SUBAPPLICATION AR_M2M_Subscribe_TO_Q_OPC (* Remote-Subscribe eines fertigen physikalischen Werts (M2M) -> VT-Anzeige (Q_NumericValue_PHYSA, gedrosselt) + VALUE_OUT. Wie AR_M2M_Subscribe_TO_Q_Publish_OPC, aber ohne lokalen Re-Publish. *)
  (* Standard: 61499-2; Description: Copyright (c) 2026 Meisterschulen am Ostbahnhof This program and the accompanying materials are made available under the terms of the Eclipse Public License 2.0 which is available at https://www.eclipse.org/legal/epl-2.0/ SPDX-License-Identifier: EPL-2.0 *)
  (* Version 1.0, 2026-10-17, Franz Höpfinger, Meisterschulen am Ostbahnhof, Kopie von AR_M2M_Subscribe_TO_Q_Publish_OPC ohne Publish/ID_WRITE (Franz: schlanke Lib-Variante bauen, damit die Lib komplett ist). Drosselung T#500ms nur auf dem Anzeige-Zweig, VALUE_OUT ungedrosselt wie im Original. *)
  PACKAGE MyLib::sys;
  IMPORT isobus::UT::Q::const::IDs::ID_NULL;
  IMPORT logiBUS::utils::conversion::phys::NumericObjectPool_S;
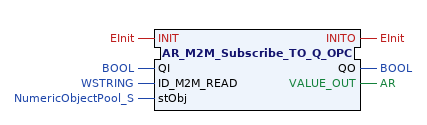
  EVENT_INPUT
    INIT : EInit; (* Initialization Request *)
  END_EVENT
  EVENT_OUTPUT
    INITO : EInit; (* Initialization Confirm *)
  END_EVENT
  VAR_INPUT
    QI : BOOL := TRUE; (* Quality Input - TRUE to enable service *)
    ID_M2M_READ : WSTRING; (* Remote-Subscribe-Adresse des fertigen physikalischen Werts (REAL) *)
    stObj : logiBUS::utils::conversion::phys::NumericObjectPool_S := (u16ObjId := ID_NULL, r32Scale := 1.0, i32Offset := 0, u8Decimals := 0); (* Object pool properties der VT-Zahlenvariable (u16ObjId, scale, offset, decimals) *)
  END_VAR
  VAR_OUTPUT
    QO : BOOL; (* Quality Output - TRUE if service executed successfully *)
  END_VAR
  PLUGS
    VALUE_OUT : adapter::types::unidirectional::AR; (* Nur-Lese-Spiegel des remote abonnierten Werts fuer weitere lokale Konsumenten *)
  END_PLUGS
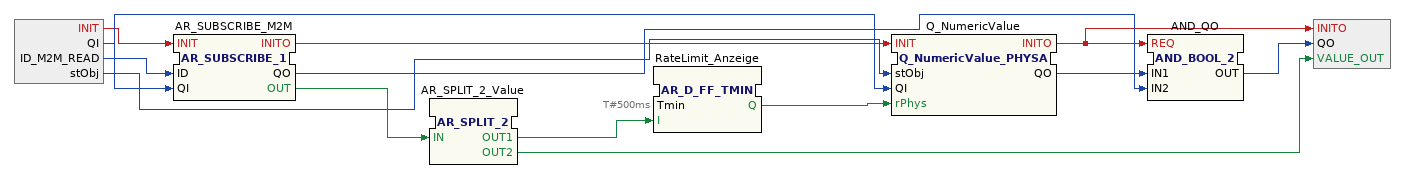
  FBS
    AR_SUBSCRIBE_M2M : adapter::net::AR_SUBSCRIBE_1;
    AR_SPLIT_2_Value : adapter::events::unidirectional::AR_SPLIT_2;
    RateLimit_Anzeige : adapter::events::unidirectional::AR_D_FF_TMIN(Tmin := T#500ms); (* Drosselt nur die VT-Anzeige auf max. 1 Update pro Tmin *)
    Q_NumericValue : isobus::UT::Q::Q_NumericValue_PHYSA;
    AND_QO : iec61131::booleanOperators::AND_BOOL_2;
  END_FBS
  EVENT_CONNECTIONS
    INIT TO AR_SUBSCRIBE_M2M.INIT;
    AR_SUBSCRIBE_M2M.INITO TO Q_NumericValue.INIT;
    Q_NumericValue.INITO TO INITO;
    Q_NumericValue.INITO TO AND_QO.REQ;
  END_CONNECTIONS
  DATA_CONNECTIONS
    ID_M2M_READ TO AR_SUBSCRIBE_M2M.ID;
    stObj TO Q_NumericValue.stObj;
    QI TO AR_SUBSCRIBE_M2M.QI;
    QI TO Q_NumericValue.QI;
    AR_SUBSCRIBE_M2M.QO TO AND_QO.IN1;
    Q_NumericValue.QO TO AND_QO.IN2;
    AND_QO.OUT TO QO;
  END_CONNECTIONS
  ADAPTER_CONNECTIONS
    AR_SUBSCRIBE_M2M.OUT TO AR_SPLIT_2_Value.IN;
    AR_SPLIT_2_Value.OUT1 TO RateLimit_Anzeige.I;
    RateLimit_Anzeige.Q TO Q_NumericValue.rPhys;
    AR_SPLIT_2_Value.OUT2 TO VALUE_OUT;
  END_CONNECTIONS
END_SUBAPPLICATION
